// TIA Portal V21 export
// export: Created 2026-11-11T00:48:16.8288122Z, ExportSetting WithDefaults, DisplayName Totally Integrated Automation Portal, DisplayVersion V21 Update 3, DisplayName STEP 7 Professional, DisplayVersion V21 Update 3, DisplayName STEP 7 Safety, DisplayVersion V21, DisplayName Tech WebApplication, DisplayVersion V21, DisplayName WinCC Basic/Comfort/Advanced, DisplayVersion V21 Update 3, DisplayName WinCC Unified, DisplayVersion V21 Update 3
FUNCTION_BLOCK "FB_Scl_sl047"   // FB187, SCL
{ S7_Optimized_Access := 'TRUE' }
VERSION : 0.1
// stored: AutoNumber true, IsIECCheckEnabled false, IsRetainMemResEnabled false, MemoryReserve 100, SetENOAutomatically false, UDAEnableTagReadback false
   VAR_INPUT
      v_in : Array[0..9] of Byte;
      v_count_in : USInt;
   END_VAR
   VAR_OUTPUT
      v_out : Array[0..9] of Bool;
   END_VAR
BEGIN
   SCATTER_BLK(IN := #v_in[0], COUNT_IN := #v_count_in, OUT => #v_out[0]);
END_FUNCTION_BLOCK
